// Communication API/CAN/CAN legacy/API/bds_can_getTxBufStatus
///This function returns the status of the Tx buffer of a CAN channel.
///
///=======
/// Remarks:
///=======
///    + Status = number of CAN messages in Tx buffer which have to be sent.
///    + The |GVL_can| is given for usage of defines.
///
///==================================================================		  			===================================================================================================
///Return value    								  									Description
///==================================================================		  			===================================================================================================
///>0																					Number of CAN messages in Tx buffer of the specified CAN channel which have to be sent.
///0																					Tx buffer is empty.
///-1																					Invalid CAN channel.
///5: BDS_CAN_FFI_ACCESS_ERROR_DU16														FFI API access error.
///
///==================================================================		   			===================================================================================================
///
///----------
/// FFI:
///----------
///This API can be used in trusted partitions. For untrusted partitions use |bds_can_getTxBufStatus_ffi|. See Freedom from Interference (FFI) concept for more details.
///
///=======
///Code Example:
///=======
///============================================================================
///
///PROGRAM appl_Task_1
///  VAR
///  
///    numMsg_s32: DINT := 16#00;
///  END_VAR
/// 
///  numMsg_s32 := bds_can_getTxBufStatus(BDS_CAN_1_D);
/// 
///  IF (numMsg_s32 > 0) THEN
///  
///    (* TX buffer contains still messages which could not be sent. If CAN channel
///       is in operational mode the messages will be sent as soon as possible. *)
///	   
///  END_IF
///END
///
///============================================================================
{attribute 'external_name' := 'cmp_rts_bds_can_getTxBufStatus'}
FUNCTION bds_can_getTxBufStatus : DINT
VAR_INPUT
	///Indicates the CAN channel.Possible values are
	///    + BDS_CAN_1_D(0)
	///    + BDS_CAN_2_D(1)
	///    + BDS_CAN_3_D(2)
	///	+ BDS_CAN_4_D(3)
	chnl_e: bds_can_Chnl_te;
END_VAR

END_FUNCTION

// Communication API/CAN/CAN_FFI_API/bds_can_getTxBufStatus_ffi
{attribute 'external_name' := 'cmp_rts_bds_can_getTxBufStatus_ffi'}
FUNCTION bds_can_getTxBufStatus_ffi : DINT
VAR_INPUT
	///Indicates the CAN channel.Possible values are
	///    + BDS_CAN_1_D(0)
	///    + BDS_CAN_2_D(1)
	///    + BDS_CAN_3_D(2)
	///	+ BDS_CAN_4_D(3)
	chnl_e: bds_can_Chnl_te;
END_VAR

END_FUNCTION

// Communication API/CAN/CAN legacy/API/bds_can_initTxDatabox
///This function initializes a CAN transmit databox.
///
///=======
/// Remarks:
///=======
///    + The use of transmit databoxes is optional!
///    + The transmit databoxes must be defined by easyConfig before using this function.
///    + Each transmit databox has to be initialized before it can be used!
///    + If a transmit databox is initialized already it can be inititalized again with new parameters. But if there is a pending message in this transmit databox it will be not sent because the databox is cleared during the initialization.
///    + The |GVL_can| is given for usage of defines.
///    + This API should be called once in Application
///
///----------
/// FFI:
///----------
///This API can be used in trusted partitions only. See Freedom from Interference (FFI) concept for more details.
///
///==================================================================		  			===================================================================================================
///Return value    								  									Description
///==================================================================		  			===================================================================================================
///0: BDS_CAN_ERR_NO_ERRORS_DU16														Function is called without errors. Transmit databox was initialized successfully.
///9: BDS_CAN_ERR_DATABOXNUM_DU16														Invalid transmit databox number.
///14: BDS_CAN_ERR_CHNL_DU16															Unknown CAN channel.
///15: BDS_CAN_ERR_ID_DU16																Invalid CAN identifier.
///16: BDS_CAN_ERR_FORMAT_DU16															Invalid message format.
///
///==================================================================		   			===================================================================================================
///
///=======
///Code Example:
///=======
///============================================================================
///
///PROGRAM PLC_PRG
///  VAR
///  	flag: BOOL;
///
///	status_u16: UINT;
///
///	DataboxData_au8: ARRAY[1..8] OF USINT;
///
///	free_count: INT;
///
///  END_VAR
///
///  (* remark: number of CAN TX databoxes must be configured in easyConfig *)
///
///  (* initialize Tx data box #1 with standard CAN Id = 16#34 *)
/// 
///IF flag = FALSE THEN
///
///	status_u16 := bds_can_initTxDatabox(BDS_CAN_1_D, 3, 16#34, BDS_CAN_STD_DU8);
///
///	bds_can_init(BDS_CAN_1_D, BDS_BAUD_500K_DU32);
///
///	flag:= TRUE;
///
///END_IF
///  (* ... *)
///END
///
///PROGRAM appl_Task_1
///  VAR
///    DataboxData_au8: ARRAY[1..8] OF USINT;
///  END_VAR
///
///  DataboxData_au8[1] := 5;
///  DataboxData_au8[2] := 7;
///
///  if (0 = bds_can_sendDatabox(BDS_CAN_3_D, 1, 2, DataboxData_au8)) THEN
///    (* ok, message will be sent. *)
///  END_IF
///END
///
///============================================================================
{attribute 'external_name' := 'cmp_rts_bds_can_initTxDatabox'}
FUNCTION bds_can_initTxDatabox : UINT
VAR_INPUT
	///Indicates the CAN channel.Possible values are
	///    + BDS_CAN_1_D(0)
	///    + BDS_CAN_2_D(1)
	///    + BDS_CAN_3_D(2)
	///	+ BDS_CAN_4_D(3)
	chnl_e: bds_can_Chnl_te;
	///Transmit databox number.
	///
	///Each transmit databox is numbered separately for each CAN channel.
	///
	///Value range: 1 .. n.
	///
	///n is the number of databoxes configured by easyConfig. 
	databoxNum_u16: UINT;
	///Identifier of CAN message.
	///
	///Value range:
	///    + 16#000 .. 16#7FF (11-bit standard format)
	///    + 16#00000000 .. 16#1FFFFFFF (29-bit extented format)
	id_u32: UDINT;
	///Indicates the format of the CAN message.
	///
	///Value range:
	///    + BDS_CAN_STD_DU8  (11-bit standard format)
	///    + BDS_CAN_EXD_DU8  (29-bit extented format)
	format_u8: USINT;
END_VAR

END_FUNCTION

// Communication API/CAN/CAN legacy/API/bds_can_sendDatabox
///Sends a message via transmit databox.
///
///=======
/// Remarks:
///=======
///    + The number of required transmit databoxes must be defined by easyConfig.
///    + The specified transmit databox has to be initialized by |bds_can_initTxDatabox| before using this function.
///    + A transmit databox buffers only the actual message.
///    + A message in a transmit databox (which was not sent) can be overwritten by a new order. No error will occur!
///    + Function |bds_can_isTxDataboxFree| can be used in order to check whether a transmit databox is free again.
///    + Messages in transmit data boxes will be sent before messages in transmit buffer (|bds_can_sendData|).
///    + The time interval for sending the messages can be defined with the function |bds_can_setTxDelay|.
///    + The |GVL_can| is given for usage of defines.
///
///----------
/// FFI:
///----------
///This API can be used in trusted partitions. For untrusted partitions use |bds_can_sendDatabox_ffi|. See Freedom from Interference (FFI) concept for more details.
///
///==================================================================		  			===================================================================================================
///Return value    								  									Description
///==================================================================		  			===================================================================================================
///0: BDS_CAN_ERR_NO_ERRORS_DU16														Function is called without errors. CAN message will be sent.
///9: BDS_CAN_ERR_DATABOXNUM_DU16														Invalid transmit databox number.
///14: BDS_CAN_ERR_CHNL_DU16															Unknown CAN channel.
///17: BDS_CAN_ERR_NUM_DATA_DU16														Invalid number of data bytes.
///60: BDS_CAN_ERR_INVALID_ADDR_DU16													Invalid address (parameter data_pau8).
///62: BDS_CAN_ERR_DATABOX_NOINIT_DU16													Transmit databox is not initialized.
///5: BDS_CAN_FFI_ACCESS_ERROR_DU16														FFI API access error.
///
///==================================================================		   			===================================================================================================
///
///=======
///Code Example:
///=======
///============================================================================
///
///PROGRAM PLC_PRG
///  VAR
///  	flag: BOOL;
///
///	status_u16: UINT;
///
///	DataboxData_au8: ARRAY[1..8] OF USINT;
///
///	free_count: INT;
///
///  END_VAR
///
///  (* remark: number of CAN TX databoxes must be configured in easyConfig *)
///
///  (* initialize Tx data box #1 with standard CAN Id = 16#34 *)
/// 
///IF flag = FALSE THEN
///
///	status_u16 := bds_can_initTxDatabox(BDS_CAN_1_D, 3, 16#34, BDS_CAN_STD_DU8);
///
///	bds_can_init(BDS_CAN_3_D, BDS_BAUD_500K_DU32);
///
///	flag:= TRUE;
///
///END_IF
///  (* ... *)
///  
///END
///
///PROGRAM appl_Task_1
///  VAR
///    DataboxData_au8: ARRAY[1..8] OF USINT;
///
///  END_VAR
///
///  DataboxData_au8[1] := 5;
///
///  DataboxData_au8[2] := 7;
///
///  if (0 = bds_can_sendDatabox(BDS_CAN_3_D, 1, 2, DataboxData_au8)) THEN
///  
///    (* ok, message will be sent. *)
///	
///  END_IF
///END
///
///============================================================================
{attribute 'external_name' := 'cmp_rts_bds_can_sendDatabox'}
FUNCTION bds_can_sendDatabox : UINT
VAR_INPUT
	///Indicates the CAN channel.Possible values are
	///    + BDS_CAN_1_D(0)
	///    + BDS_CAN_2_D(1)
	///    + BDS_CAN_3_D(2)
	///	+ BDS_CAN_4_D(3)
	chnl_e: bds_can_Chnl_te;
	///Transmit databox number.
	///
	///Each transmit databox is numbered separately for each CAN channel.
	///
	///Value range: 1 .. n.
	///
	///n is the number of Tx databoxes configured by easyConfig. 
	txDataboxNum_u16: UINT;
	///Number of bytes to be sent.
	///
	///Value range: 0 .. 8
	numBytes_u8: USINT;
	///Pointer to array of data bytes. The number of bytes is contained in parameter numBytes_u8. A NULL pointer is allowed if number of data bytes (parameter numBytes_u8) is zero. 
	data_pau8: POINTER TO USINT;
END_VAR

END_FUNCTION

// Communication API/CAN/CAN legacy/API/bds_can_isTxDataboxFree
///This function checks whether a transmit databox is free again. A transmit databox is free again if it was possible to send the last CAN message via the bus.
///
///=======
/// Remarks:
///=======
///    + The use of transmit databoxes is optional!
///    + The transmit databoxes of that CAN channel has to be defined by easyConfig tool and that transmit databox has to be initialised by bds_can_initTxDatabox before using this function.
///    + This function can be used to prevent overwriting of a message that has not yet been sent in a send databox, by checking whether the previous message was actually sent before writing the new message to the databox.
///    + How quickly a databox is free again for sending greatly depends on the baud rate and the bus load.
///    + The |GVL_can| is given for usage of defines.
///
///----------
/// FFI:
///----------
///This API can be used in trusted partitions. For untrusted partitions use |bds_can_isTxChannelFree_ffi|. See Freedom from Interference (FFI) concept for more details.
///
///==================================================================		  			===================================================================================================
///Return value    								  									Description
///==================================================================		  			===================================================================================================
///0: BDS_CAN_TX_DATABOX_EMPTY_DU16													No error. Databox is empty.
///1: BDS_CAN_TX_DATABOX_NOT_EMPTY_DU16												No error. Databox is not empty.
///9: BDS_CAN_ERR_DATABOXNUM_DU16														Invalid databox number.
///14: BDS_CAN_ERR_CHNL_DU16															Unknown CAN channel.
///62: BDS_CAN_ERR_DATABOX_NOINIT_DU16													Databox is not initialized.
///5: BDS_CAN_FFI_ACCESS_ERROR_DU16														FFI API access error.
///
///==================================================================		   			===================================================================================================
///
///=======
///Code Example:
///=======
///============================================================================
///
///PROGRAM PLC_PRG
///
///  VAR
///  	flag: BOOL;
///
///	status_u16: UINT;
///
///	DataboxData_au8: ARRAY[1..8] OF USINT;
///
///	free_count: INT;
///
///  END_VAR
///
///  (* remark: number of CAN TX databoxes must be configured in easyConfig *)
///
///  (* initialize Tx data box #1 with standard CAN Id = 16#34 *)
/// 
///IF flag = FALSE THEN
///
///	status_u16 := bds_can_initTxDatabox(BDS_CAN_1_D, 3, 16#34, BDS_CAN_STD_DU8);
///
///	bds_can_init(BDS_CAN_1_D, BDS_BAUD_500K_DU32);
///
///	flag:= TRUE;
///
///END_IF
///
///PROGRAM appl_Task_1
///  VAR
///  
///  END_VAR
///
///  IF (0 = bds_can_isTxDataboxFree(BDS_CAN_1_D, 1)) THEN
///  
///    (* transmit databox 1 on CAN channel 1 is free and can be loaded again *)
///    (* ... *)
///	
///  END_IF
///END
///
///============================================================================
{attribute 'external_name' := 'cmp_rts_bds_can_isTxDataboxFree'}
FUNCTION bds_can_isTxDataboxFree : UINT
VAR_INPUT
	///Indicates the CAN channel.Possible values are
	///    + BDS_CAN_1_D(0)
	///    + BDS_CAN_2_D(1)
	///    + BDS_CAN_3_D(2)
	///	+ BDS_CAN_4_D(3)
	chnl_e: bds_can_Chnl_te;
	///Transmit databox number.
	///
	///Each transmit databox is numbered separately for each CAN channel.
	///
	///Value range: 1 .. n.
	///
	///n is the number of databoxes configured by easyConfig. 
	txDataboxNum_u16: UINT;
END_VAR

END_FUNCTION

// Communication API/CAN/CAN_FFI_API/bds_can_isTxChannelFree_ffi
{attribute 'external_name' := 'cmp_rts_bds_can_isTxChannelFree_ffi'}
FUNCTION bds_can_isTxChannelFree_ffi : UINT
VAR_INPUT
	///Indicates the CAN channel.Possible values are
	///    + BDS_CAN_1_D(0)
	///    + BDS_CAN_2_D(1)
	///    + BDS_CAN_3_D(2)
	///	+ BDS_CAN_4_D(3)
	chnl_e: bds_can_Chnl_te;
END_VAR

END_FUNCTION

// Communication API/CAN/CAN legacy/API/bds_can_sendData
///Sends a message via the specified CAN channel.
///
///=======
/// Remarks:
///=======
///    + The CAN channel is not buffered until a buffer is registered within easyConfig.
///    + If a buffer is registered then messages are saved in buffer and will be sent in a background process as fast as possible. The buffer principle is first in first out (FIFO).
///    + The time interval for sending the messages can be defined with the function |bds_can_setTxDelay|.
///    + Messages in transmit data boxes (|bds_can_sendDatabox|) will be sent before messages in transmit buffer (|bds_can_sendData|).
///    + The |GVL_can| is given for usage of defines.
///
///----------
/// FFI:
///----------
///This API can be used in trusted partitions. For untrusted partitions use |bds_can_sendData_ffi|. See Freedom from Interference (FFI) concept for more details.
///
///==================================================================		  			===================================================================================================
///Return value    								  									Description
///==================================================================		  			===================================================================================================
///0: BDS_CAN_ERR_NO_ERRORS_DU16														Function is called without errors. CAN message will be sent.
///14: BDS_CAN_ERR_CHNL_DU16															Unknown CAN channel.
///15: BDS_CAN_ERR_ID_DU16																Invalid CAN identifier.
///16: BDS_CAN_ERR_FORMAT_DU16															Invalid message format.
///17: BDS_CAN_ERR_NUM_DATA_DU16														Invalid number of data bytes.
///20: BDS_CAN_ERR_TXBUF_OVFL_DU16														CAN message could not be sent, because of send buffer is full. *1)
///60: BDS_CAN_ERR_INVALID_ADDR_DU16													Invalid address (parameter data_pau8).
///5: BDS_CAN_FFI_ACCESS_ERROR_DU16														FFI API access error.
///
///==================================================================		   			===================================================================================================
///
///possible reasons:
///    + API
///	    + No can send buffer was registered or buffer registered is too small; see buffer configuration in easyConfig.
///        + To many CAN messages have to be sent per time (more orders exceed performance of sending); use higher baudrate, see bds_can_init()
///        + To many CAN messages have to be sent per time by CAN send databoxes; (sending by databoxes is preferred! see bds_can_sendDatabox()
///        + A TX delay time with bds_can_setTxDelay() is defined, which is too big for the number of messages to be sent.
///    + External factors
///        + CAN bus is busy by CAN messages with higher priorities sending by other ECU's so that CAN messages of the own ECU can not be sent.
///        + The sending of CAN messages is delayed due to CAN BUS error(s). Bus-off states will be recovered automatically.
///
///=======
///Code Example:
///=======
///============================================================================
///
///PROGRAM PLC_PRG
///  VAR
///  
///  END_VAR
///
///  (* remark: a CAN TX buffer must be configured in easyConfig *)
///
///  (* re-initialize can channel 1 with 250KBaud. Call the bds_can_init API once *)
///  
///  bds_can_init(BDS_CAN_1_D, BDS_BAUD_250K_DU32);
///
///  (* ... *)
///  
///END
///
///PROGRAM appl_Task_1
///  VAR
///    data_au8: ARRAY[0..7] OF USINT;
///  END_VAR
///
///  data_au8[0] := 5;
///  data_au8[1] := 7;
///
///  IF (0 = bds_can_sendData(BDS_CAN_1_D, 16#123456, BDS_CAN_EXD_DU8, 2, ADR(data_au8))) THEN
///  
///    (* ok, message is buffered and will be sent as fast as possible. *)
///	
///  END_IF
///END
///
///============================================================================
{attribute 'external_name' := 'cmp_rts_bds_can_sendData'}
FUNCTION bds_can_sendData : UINT
VAR_INPUT
	///Indicates the CAN channel.Possible values are
	///    + BDS_CAN_1_D(0)
	///    + BDS_CAN_2_D(1)
	///    + BDS_CAN_3_D(2)
	///	+ BDS_CAN_4_D(3)
	chnl_e: bds_can_Chnl_te;
	///Identifier of CAN message.
	///
	///Value range:
	///    - 16#000 .. 16#7FF (11-bit standard format)
	///    - 16#00000000 .. 16#1FFFFFFF (29-bit extented format)
	id_u32: UDINT;
	///Indicates the format of the CAN message.
	///
	///Value range:
	///    + BDS_CAN_STD_DU8  (11-bit standard format)
	///    + BDS_CAN_EXD_DU8  (29-bit extented format)
	format_u8: USINT;
	///Number of bytes to be sent.
	///
	///Value range: 0 .. 8
	numBytes_u8: USINT;
	///Pointer to array of data bytes. The number of bytes is contained in parameter numBytes_u8. A NULL pointer is allowed if number of data bytes (parameter numBytes_u8) is zero. 
	data_pau8: POINTER TO USINT;
END_VAR

END_FUNCTION

// Communication API/CAN/CAN legacy/API/bds_can_setTxDelay
///The bds_can_setTxDelay function can be used to define an optional delay time for sending CAN messages.
///
///=======
/// Remarks:
///=======
///    + Without executing this function the default delay time = 0 is used.
///    + A delay time > 0 should be only specified, if another controller is not able to receive the CAN messages with full speed.
///    + For each CAN channel another delay time can be specified.
///    + Only messages which are sent with the functions |bds_can_sendDatabox|, |bds_can_sendData| and all messages of ISOBUS module will be delayed.
///    + Signal based CAN messages, XCP and UDS messages are not impacted by this function.
///    + If an error occurs during execution of this function, the actual delay time will be not modified.
///    + The |GVL_can| is given for usage of defines.
///
///----------
/// FFI:
///----------
///This API can be used in trusted partitions only. See Freedom from Interference (FFI) concept for more details.
///
///==================================================================		  			===================================================================================================
///Return value    								  									Description
///==================================================================		  			===================================================================================================
///0: BDS_CAN_ERR_NO_ERRORS_DU16														Function is called without errors. Message data returned in msg_s are valid.
///14: BDS_CAN_ERR_CHNL_DU16															Unknown CAN channel.
///
///==================================================================		   			===================================================================================================
///
///=======
///Code Example:
///=======
///============================================================================
///
///PROGRAM PLC_PRG
///  VAR
///  
///  END_VAR
///
///  (* set the minimum TX delay time to 2ms for CAN channel 1 *)
///  
///IF flag = FALSE THEN
///
///	  bds_can_setTxDelay(BDS_CAN_1_D, 2);
///
///	flag:= TRUE;
///
///END_IF
///  (* ... *)
///END
///
///============================================================================
{attribute 'external_name' := 'cmp_rts_bds_can_setTxDelay'}
FUNCTION bds_can_setTxDelay : UINT
VAR_INPUT
	///Indicates the CAN channel.Possible values are
	///    + BDS_CAN_1_D(0)
	///    + BDS_CAN_2_D(1)
	///    + BDS_CAN_3_D(2)
	///	+ BDS_CAN_4_D(3)
	chnl_e: bds_can_Chnl_te;
	///Minimum delay time in ms between two sent can messages.
	///
	///Value range: 0 .. 65535.
	///
	///0 = no delay time, means that the can messages will be sent as fast as possible.
	time_u16: UINT;
END_VAR

END_FUNCTION

// Communication API/CAN/CAN_FFI_API/bds_can_sendData_ffi
{attribute 'external_name' := 'cmp_rts_bds_can_sendData_ffi'}
FUNCTION bds_can_sendData_ffi : UINT
VAR_INPUT
	///Indicates the CAN channel.Possible values are
	///    + BDS_CAN_1_D(0)
	///    + BDS_CAN_2_D(1)
	///    + BDS_CAN_3_D(2)
	///	+ BDS_CAN_4_D(3)
	chnl_e: bds_can_Chnl_te;
	///Identifier of CAN message.
	///
	///Value range:
	///    - 16#000 .. 16#7FF (11-bit standard format)
	///    - 16#00000000 .. 16#1FFFFFFF (29-bit extented format)
	id_u32: UDINT;
	///Indicates the format of the CAN message.
	///
	///Value range:
	///    + BDS_CAN_STD_DU8  (11-bit standard format)
	///    + BDS_CAN_EXD_DU8  (29-bit extented format)
	format_u8: USINT;
	///Number of bytes to be sent.
	///
	///Value range: 0 .. 8
	numBytes_u8: USINT;
	///Pointer to array of data bytes. The number of bytes is contained in parameter numBytes_u8. A NULL pointer is allowed if number of data bytes (parameter numBytes_u8) is zero. 
	data_pau8: POINTER TO USINT;
END_VAR

END_FUNCTION

// Communication API/CAN/CAN_FFI_API/bds_can_sendDatabox_ffi
{attribute 'external_name' := 'cmp_rts_bds_can_sendDatabox_ffi'}
FUNCTION bds_can_sendDatabox_ffi : UINT
VAR_INPUT
	///Indicates the CAN channel.Possible values are
	///    + BDS_CAN_1_D(0)
	///    + BDS_CAN_2_D(1)
	///    + BDS_CAN_3_D(2)
	///	+ BDS_CAN_4_D(3)
	chnl_e: bds_can_Chnl_te;
	///Transmit databox number.
	///
	///Each transmit databox is numbered separately for each CAN channel.
	///
	///Value range: 1 .. n.
	///
	///n is the number of Tx databoxes configured by easyConfig. 
	txDataboxNum_u16: UINT;
	///Number of bytes to be sent.
	///
	///Value range: 0 .. 8
	numBytes_u8: USINT;
	///Pointer to array of data bytes. The number of bytes is contained in parameter numBytes_u8. A NULL pointer is allowed if number of data bytes (parameter numBytes_u8) is zero. 
	data_pau8: POINTER TO USINT;
END_VAR

END_FUNCTION

// Communication API/CAN/CAN legacy/API/bds_can_isTxChannelFree
///This function checks whether a complete CAN transmit channel is empty.
///
///=======
/// Remarks:
///=======
///    + Empty means that there is no message to send in hardware CAN controller and in any Tx databox (if registered and initialized) and Tx buffer (if registered) is empty.
///    + This function can be used in order to check if a previous message was sent completely on CAN bus. 
///    + The |GVL_can| is given for usage of defines.
///
///----------
/// FFI:
///----------
///This API can be used in trusted partitions. For untrusted partitions use |bds_can_isTxDataboxFree_ffi|. See Freedom from Interference (FFI) concept for more details.
///
///==================================================================		  			===================================================================================================
///Return value    								  									Description
///==================================================================		  			===================================================================================================
///0: BDS_CAN_TX_CHANNEL_EMPTY_DU16													No error. CAN transmit channel is empty. No CAN message has to be sent at the moment.
///1: BDS_CAN_TX_CHANNEL_NOT_EMPTY_DU16												No error. CAN transmit channel is not empty. Sending of a message is still in progress and/or CAN Tx messages are still buffered for sending. 
///2: BDS_CAN_TX_CHANNEL_INV_CAN_DU16													Unknown CAN channel.
///5: BDS_CAN_FFI_ACCESS_ERROR_DU16														FFI API access error.
///
///==================================================================		   			===================================================================================================
///
///=======
///Code Example:
///=======
///============================================================================
///
///PROGRAM appl_Task_1
///  VAR
///  
///  END_VAR
///
///  IF (BDS_CAN_TX_CHANNEL_EMPTY_DU16 = bds_can_isTxChannelFree(BDS_CAN_1_D)) THEN
///  
///    (* All TX databoxes and TX buffer on CAN channel 1 are empty. *)
///    (* ... *)
///	
///  END_IF
///END
///
///============================================================================
{attribute 'external_name' := 'cmp_rts_bds_can_isTxChannelFree'}
FUNCTION bds_can_isTxChannelFree : UINT
VAR_INPUT
	///Indicates the CAN channel.Possible values are
	///    + BDS_CAN_1_D(0)
	///    + BDS_CAN_2_D(1)
	///    + BDS_CAN_3_D(2)
	///	+ BDS_CAN_4_D(3)
	chnl_e: bds_can_Chnl_te;
END_VAR

END_FUNCTION

// Communication API/CAN/CAN_FFI_API/bds_can_isTxDataboxFree_ffi
{attribute 'external_name' := 'cmp_rts_bds_can_isTxDataboxFree_ffi'}
FUNCTION bds_can_isTxDataboxFree_ffi : UINT
VAR_INPUT
	///Indicates the CAN channel.Possible values are
	///    + BDS_CAN_1_D(0)
	///    + BDS_CAN_2_D(1)
	///    + BDS_CAN_3_D(2)
	///	+ BDS_CAN_4_D(3)
	chnl_e: bds_can_Chnl_te;
	///Transmit databox number.
	///
	///Each transmit databox is numbered separately for each CAN channel.
	///
	///Value range: 1 .. n.
	///
	///n is the number of databoxes configured by easyConfig. 
	txDataboxNum_u16: UINT;
END_VAR

END_FUNCTION

// Communication API/CAN/CAN signal based/API/bds_can_sendSignal
///This function is used to transmit message with signal data specified by signal ID on the CAN bus.
///
///Signals are part of PDU, call to this API would cause the PDU to be sent on bus but with the signal contents updated by the signal data pointer. 
///
///This API is responsible for transmission of PDU (for Tx mode= Direct) and updation of signal data (for Tx mode= Cyclic).
///
///=======
/// Remarks:
///=======
///    + Signals referred here are available upon a valid DBC import. 
///    + The parameters of the signal such as Signal ID, length and signal data pointer are passed as parameters to the function while the CAN ID would correspond to the PDU the signal is mapped to.
///    + Easy Config tool allows import of DBC file and selection of frames and signals for the respective CAN nodes.
///    + Signal and PDU properties like Transmission type, no. of repetitions, signal length and so on shall be configured from easyConfig cloud tool.
///    + Interaction Layer Protocol Data Unit(IPDU - a collection of messages transmitted between nodes in a network. 
///    + A sending node packs the messages into an I-PDU in the Interaction Layer (IL) and then transmits them to the network in the Data Link Layer (DLL). 
///    + A receiving node passes each I-PDU from the DLL and to the IL. There, it unpacks the messages and use their contents in the application.
///    + The |GVL_can| is given for usage of defines.
///    + Signal IDs can be located in the post build configuration file - linCanSignals_easyConfig.xml.
///
///----------
/// FFI:
///----------
///This API can be used in trusted partitions only. See Freedom from Interference (FFI) concept for more details.
///
///----------
/// NOTICE:
///----------
///- For signals imported from dbc file,the signal type information comes from dbc. This would generally be of static types like USINT, UINT, SINT, INT. In order to be able to change the length of signal, it requires that the signal is of type USINT_DYN.
///So, for all signals imported from dbc, the length parameter in API has to be set to 0.
///
///==================================================================		  			===================================================================================================
///Return value    								  									Description
///==================================================================		  			===================================================================================================
///BDS_CAN_ERR_NO_ERRORS_DU16 (= 0)													Signal transmission successful.
///BDS_CANSIG_ERR_TX_FAIL_DU16(=117)													Transmission failure.
///BDS_CANSIG_ERR_TX_NOSERVICE_DU16(=119)												Service not available-PDU inactive.
///BDS_CANSIG_ERR_TX_DATAPTR_DU16(=114)												Invalid data pointer address.
///BDS_CANSIG_ERR_NUM_TX_SIG_DU16(=112)												Invalid Signal ID.
///
///==================================================================		   			===================================================================================================
///
///=======
///Code Example:
///=======
///============================================================================
///
///PROGRAM appl_10ms_task
///  VAR
///  
///    bds_IPduGrpVctr_au8:ARRAY[0..1] OF USINT;
///	
///    signaldata_au8: ARRAY[0..7] OF USINT;
///	
///    length_u16: UINT := 16#00;
///	
///  END_VAR
///
///   (* Set the I-PDU and corresponding groups *)
///   (* PDU ,signal and group Ids are available in post build config files from easyConfig *)
/// 
///   bds_can_setMsgGroup(ADR(bds_IPduGrpVctr_au8),ComConf_ComIPduGroup_ComIPduGroup_C_Tx, 1);
///   
///   bds_can_startAllMsgGroups(ADR(bds_IPduGrpVctr_au8), 1) ;
///
///   IF ( 0 = bds_can_sendSignal(ComConf_ComSignal_ComSignal_C_xTx, ADR(signaldata_au8), length_u16) ) THEN
///   
///     (* ok,message is sent on bus with updated signal data *)
///   END_IF
///END
///
///============================================================================
{attribute 'external_name' := 'cmp_rts_bds_can_sendSignal'}
FUNCTION bds_can_sendSignal : UINT
VAR_INPUT
	///ID of the signal to be sent.
	signalId_u16: UINT;
	///Pointer array to the data to be transmitted.
	signalDataPtr_au8: POINTER TO USINT;
	///No. of bytes of data to be sent (for dynamic type signal)
	///	
	///- 0, for static type signals (imported from dbc, refer NOTICE above)
	length_u16: UINT;
END_VAR

END_FUNCTION

// Communication API/CAN/CAN signal based/API/bds_can_setMsgGroup
///A PDU group contains multiple PDUs and each PDU contains one or more signals.
///
///Every message/PDU should be activated before communication. To do this it is required to activate the PDU group in which it is present. This function sets the PDU group specified by group ID, which has to be enabled later by API |bds_can_startAllMsgGroups|.
///
///   
///=======
/// Remarks:
///=======
///    + PDU and message are the same in this context. When it is said that PDU is active, it also means that the message is active.
///    + PDUs referred here are available upon a valid DBC import. 
///    + With the available resources of RC18-12/40 and RC27-18/40, PDU group: There can be a maximum of 8 PDU groups based on the 4 CAN nodes and for each direction (transmit/receive). When PDUs are imported into CAN nodes on eC by DBC importer, the PDUs are put into respective groups. 
///    + To set a PDU, it is necessary to set the PDU group that contains the PDU. 
///    + This API can be called anywhere in the ASW - at init or inside cyclic task.
///    + The PDU groups are generated when we import DBC or add the frame to the CAN channel from eC.
///    + The PDU group name generated will look like ComConf_ComIPduGroup_ComIPduGroup_CAN "channel number"_TX and  ComConf_ComIPduGroup_ComIPduGroup_CAN "channel number"_RX. 
///    + Example:  For CAN 3 the PDU group will look like "ComConf_ComIPduGroup_ComIPduGroup_CAN_3_TX" and   "ComConf_ComIPduGroup_ComIPduGroup_CAN_3_RX".
///    + Interaction Layer Protocol Data Unit (IPDU) - a collection of messages transmitted between nodes in a network. 
///    + A sending node packs the messages into an I-PDU in the Interaction Layer (IL) and then transmits them to the network in the Data Link Layer (DLL). 
///    + A receiving node passes each I-PDU from the DLL and to the IL. There, it unpacks the messages and use their contents in the application.
///	   + The |GVL_can| is given for usage of defines.
///    + PDU and PDU group IDs can be located in the post build configuration file - linCanSignals_easyConfig.xml.
///
///----------
/// FFI:
///----------
///This API can be used in trusted partitions only. See Freedom from Interference (FFI) concept for more details.
///
///==================================================================		  			===================================================================================================
///Return value    								  									Description
///==================================================================		  			===================================================================================================
///BDS_CAN_ERR_NO_ERRORS_DU16 (= 0)													PDU group setting successful.
///BDS_CANSIG_ERR_NULLIPDUVECTOR_DU16(=110)											Invalid Group vector array address.
///BDS_CANSIG_ERR_BITFLAG_DU16(=111)													Invalid parameter bitval.
///
///==================================================================		   			===================================================================================================
///
///=======
///Code Example:
///=======
///============================================================================
///
///PROGRAM appl_10ms_task
///  VAR
///  
///    bds_IPduGrpVctr_au8:ARRAY[0..1] OF USINT;
///  END_VAR
///
///IF ( 0 = bds_can_setMsgGroup(ADR(bds_IPduGrpVctr_au8),ComConf_ComIPduGroup_ComIPduGroup_CAN_1_Tx, 1) ) THEN
///
///    (* ComIPduGroup_CAN_1_TX PDU group is set successfully *)
///    (* All PDUs of this group is now set, next step is to enable *)
///END_IF
///END
///
///============================================================================
{attribute 'external_name' := 'cmp_rts_bds_can_setMsgGroup'}
FUNCTION bds_can_setMsgGroup : UINT
VAR_INPUT
	///PDU group array containing the activation state (stopped = 0/ started = 1) for all message groups.
	rbr_iPduGrpVctr_au8: POINTER TO ARRAY[0..1] OF USINT;
	///PDU group used to identify the corresponding bit in the message group vector.
	ipduGroupId_u16: UINT;
	///New value of the corresponding bit(set PDU =1; reset PDU=0).
	bitval_u8: USINT;
END_VAR

END_FUNCTION

// Communication API/CAN/CAN signal based/API/bds_can_startAllMsgGroups
///This is the master function responsible for activating or deactivating PDU/message groups.
///
///This function is used to activate all PDU/message groups that were set by |bds_can_setMsgGroup|. 
///
///When a PDU group is activated by means of call to this API, all the PDUs belonging to these groups would be activated and the contained signals would be ready for transmission or reception.
///
///=======
/// Remarks:
///=======
///    + PDU and message are the same in this context. 
///    + PDUs referred here are available upon a valid DBC import. 
///    + It is sufficient to call this API once after setting all the PDU groups using the API  |bds_can_setMsgGroup|.
///    + If suppose |bds_can_setMsgGroup| is called sometime later after |bds_can_startAllMsgGroups|, the new PDU group set is still not active and so, bds_can_startAllMsgGroups() will have to be called again. So, everytime a new PDU group is set, it should be activated with this API.
///    + For cyclic signals, the transmission will start soon after the corresponding message and message group is activated by call to this API, the signal data at this instant would be the signal init value defined in eC. Signal data gets updated when the API |bds_can_sendSignal| is called later.
///    + For direct signals, transmission will happen only upon call to |bds_can_sendSignal|.
///    + Interaction Layer Protocol Data Unit(IPDU) - a collection of messages transmitted between nodes in a network. 
///    + A sending node packs the messages into an I-PDU in the Interaction Layer (IL) and then transmits them to the network in the Data Link Layer (DLL). 
///    + A receiving node passes each I-PDU from the DLL and to the IL. There, it unpacks the messages and use their contents in the application.
///    + The |GVL_can| is given for usage of defines.
///    + PDU and PDU group IDs can be located in the post build configuration file - linCanSignals_easyConfig.xml.
///
///----------
/// FFI:
///----------
///This API can be used in trusted partitions only. See Freedom from Interference (FFI) concept for more details.
///
///==================================================================		  			===================================================================================================
///Return value    								  									Description
///==================================================================		  			===================================================================================================
///BDS_CAN_ERR_NO_ERRORS_DU16 (= 0)													PDU groups activation successful.
///BDS_CANSIG_ERR_NULLIPDUVECTOR_DU16(=110)											Invalid Group vector array address.
///BDS_CANSIG_ERR_BITFLAG_DU16(=111)													Invalid parameter Initialize.
///
///==================================================================		   			===================================================================================================
///
///=======
///Code Example:
///=======
///============================================================================
///
///PROGRAM appl_task_1
///  VAR
///  
///    bds_IPduGrpVctr_au8:ARRAY[0..1] OF USINT;
///  END_VAR
///
///bds_can_setMsgGroup(ADR(bds_IPduGrpVctr_au8),ComConf_ComIPduGroup_ComIPduGroup_CAN_1_Tx, 1);
///
///IF ( 0 = bds_can_startAllMsgGroups(ADR(bds_IPduGrpVctr_au8), 1) ) THEN
///
///  (* PDU groups are active and signals ready for transmission(direct) or signal transmission started(cyclic) *)
///END_IF
///END
///
///============================================================================
{attribute 'external_name' := 'cmp_rts_bds_can_startAllMsgGroups'}
FUNCTION bds_can_startAllMsgGroups : UINT
VAR_INPUT
	///PDU group array containing the activation state (stopped = 0/ started = 1) for all PDU groups.
	rbr_iPduGrpVctr_au8: POINTER TO ARRAY[0..1] OF USINT;
	///flag to request initialization of the PDUs
	///	
	///0 = PDU groups will not be activated
	///
	///1 = PDU groups will be activated
	initialize_u8: USINT;
END_VAR

END_FUNCTION

// Communication API/CAN/CAN signal based/API/bds_can_sendSignalGroup
///This function sends the signal group data on the PDU/message.
///
///=======
/// Remarks:
///=======
///    + Before call to this API, it is necessary to update the signal group with data for every group signal belonging to signal group. This is done by using the API bds_can_setGroupSignalData. This function then sends the contents of shadow buffer on the PDU.
///    + Group signals and Signal groups referred here are available upon a valid DBC import. 
///    + Additionally, modification of signal groups by adding group signals to signal group can be done on easyConfig cloud tool.
///    + The parameter SignalGroup ID is passed as parameter to the function while the CAN ID would correspond to the PDU the signal group is mapped to.
///    + Cloud tool allows import of DBC file and selection of frames and signals for the respective CAN nodes.
///    + Signal and PDU properties like Transmission type, number of repetitions, signal length and so on shall be configured from easyConfig cloud tool.
///    + Interaction Layer Protocol Data Unit (IPDU - a collection of messages transmitted between nodes in a network). 
///    + A sending node packs the messages into an I-PDU in the Interaction Layer (IL) and then transmits them to the network in the Data Link Layer (DLL). 
///    + A receiving node passes each I-PDU from the DLL and to the IL. There, it unpacks the messages and use their contents in the application.
///    + The |GVL_can| is given for usage of defines.
///    + Group Signal IDs can be located in the post build configuration file - linCanSignals_easyConfig.xml.
///
///----------
/// FFI:
///----------
///This API can be used in trusted partitions only. See Freedom from Interference (FFI) concept for more details.
///
///==================================================================		  			===================================================================================================
///Return value    								  									Description
///==================================================================		  			===================================================================================================
///BDS_CAN_ERR_NO_ERRORS_DU16 (= 0)													Transmission successful.
///BDS_CANSIG_ERR_TX_NOSERVICE_DU16(=119)												Service not available-PDU inactive.
///
///==================================================================		   			===================================================================================================
///
///=======
///Code Example:
///=======
///============================================================================
///
///PROGRAM appl_task_1
///  VAR
///  
///    bds_IPduGrpVctr_au8:ARRAY[0..1] OF USINT;
///	
///    signaldata_u64: ULINT := 16#1234;
///  END_VAR
///
///  (* Set the I-PDU and corresponding groups *)
///  (* PDU ,signal and group Ids are available in post build config files from easyConfig *)
/// 
///   bds_can_setMsgGroup(ADR(bds_IPduGrpVctr_au8),ComConf_ComIPduGroup_ComIPduGroup_C_Tx, 1);
///   
///   bds_can_startAllMsgGroups(ADR(bds_IPduGrpVctr_au8), 1) ;
///
///   (* update group signal data *)
///   
///   bds_can_setGroupSignalData(ComConf_ComGroupSignal_ComGroupSignal_Tx, signaldata_u64);
///
///   IF ( 0 = bds_can_sendSignalGroup(ComConf_ComSignalGroup_ComSignalGroup_Tx_1) ) THEN
///   
///     (* ok, message is sent on bus with signalgroup data *)
///   END_IF
///END
///
///============================================================================
{attribute 'external_name' := 'cmp_rts_bds_can_sendSignalGroup'}
FUNCTION bds_can_sendSignalGroup : UINT
VAR_INPUT
	///ID of the signal group to be transmitted.
	signalGroupId_u16: UINT;
END_VAR

END_FUNCTION

// Communication API/CAN/CAN signal based/API/bds_can_setGroupSignalData
///This function updates the group signal with the data referenced by signalData parameter.
///
///The updated data is now stored in a shadow buffer of the signal group.
///
///The entire contents of signal group shadow buffer is transmitted on a message/PDU upon call to API |bds_can_sendSignalGroup|.
///
///=======
/// Remarks:
///=======
///    + Group Signals and Signal groups referred here are available upon a valid DBC import. 
///    + Additionally, modification of signal groups by adding group signals to signal group can be done on easyConfig cloud tool.
///    + Group Signal IDs can be located in the post build configuration file - BODAS API library, bds_rts_ec.xml.
///    + The parameters of the signal such as Group Signal ID and signal data are passed as parameters to the function while the CAN ID would correspond to. 
///    + Interaction Layer Protocol Data Unit (IPDU - a collection of messages transmitted between nodes in a network). 
///    + A sending node packs the messages into an I-PDU in the Interaction Layer (IL) and then transmits them to the network in the Data Link Layer (DLL). 
///    + A receiving node passes each I-PDU from the DLL and to the IL. There, it unpacks the messages and use their contents in the application.
///    + The |GVL_can| is given for usage of defines.
///    + Group Signal IDs can be located in the post build configuration file - linCanSignals_easyConfig.xml.
///
///----------
/// FFI:
///----------
///This API can be used in trusted partitions only. See Freedom from Interference (FFI) concept for more details.
///
///==================================================================		  			===================================================================================================
///Parameter	   								  										Description
///==================================================================		  			===================================================================================================
///groupSignalId_u16																	ID of the group signal to be sent.
///signalData_u64																		Signal data for the specified group signal to be transmitted. Maximum size of data is 64 bits(8bytes).
///
///==================================================================		   			===================================================================================================
///
///=======
///Code Example:
///=======
///============================================================================
///
///PROGRAM appl_10ms_task
///  VAR
///  
///    bds_IPduGrpVctr_au8:ARRAY[0..1] OF USINT;
///	
///    signaldata_u64: ULINT := 16#1234;
///  END_VAR
///
///  (* Set the I-PDU and corresponding groups *)
///  (* PDU ,signal and group Ids are available in post build config files from easyConfig *)
/// 
///   bds_can_setMsgGroup(ADR(bds_IPduGrpVctr_au8),ComConf_ComIPduGroup_ComIPduGroup_C_Tx, 1);
///   
///   bds_can_startAllMsgGroups(ADR(bds_IPduGrpVctr_au8), 1) ;
///
///   (* update group signal data *)
///   
///   bds_can_setGroupSignalData(ComConf_ComGroupSignal_ComGroupSignal_Tx, signaldata_u64);
///END
///
///============================================================================
{attribute 'external_name' := 'cmp_rts_bds_can_setGroupSignalData'}
FUNCTION bds_can_setGroupSignalData : BOOL
VAR_INPUT
	///ID of the group signal to be sent.
	groupSignalId_u16: UINT;
	///Signal data for the specified group signal to be transmitted. Maximum size of data is 64 bits(8bytes).
	signalData_u64: ULINT;
END_VAR

END_FUNCTION

// Communication API/CAN/CAN signal based/API/bds_can_receiveSignal
///Signals are part of PDU/message, call to this API would cause the signal data of the PDU/message received on bus to be copied to application defined buffer.
///
///=======
/// Remarks:
///=======
///    + Signals referred here are available upon a valid DBC import. 
///    + The parameters of the signal such as Signal ID, length and signal data pointer are passed as parameters to the function while the CAN ID would correspond to the PDU, the signal is mapped to.
///    + Easy Config tool allows import of DBC file and selection of frames and signals for the respective CAN nodes.
///    + Signal and PDU properties like Transmission type, no. of repetitions, signal length and so on shall be configured from easyConfig cloud tool.
///    + Interaction Layer Protocol Data Unit (IPDU - a collection of messages transmitted between nodes in a network). 
///    + A sending node packs the messages into an I-PDU in the Interaction Layer (IL) and then transmits them to the network in the Data Link Layer (DLL). 
///    + A receiving node passes each I-PDU from the DLL and to the IL. There, it unpacks the messages and use their contents in the application.
///    + The |GVL_can| is given for usage of defines.
///    + Signal IDs can be located in the post build configuration file - linCanSignals_easyConfig.xml.
///
///----------
/// FFI:
///----------
///This API can be used in trusted partitions only. See Freedom from Interference (FFI) concept for more details.
///
///----------
/// NOTICE:
///----------
///The length parameter specifies the no. of bytes of data to be received and it is important to specify exactly the no. of incoming bytes else it would result in length validation failure.
///- For signals imported from dbc file,the signal type information comes from dbc. This would generally be of static types like USINT, UINT, SINT, INT.
///
///==================================================================		  			===================================================================================================
///Return value    								  									Description
///==================================================================		  			===================================================================================================
///BDS_CAN_ERR_NO_ERRORS_DU16 (= 0)													Signal reception successful.
///BDS_CANSIG_ERR_RX_FAIL_DU16(=118)													Reception failure.
///BDS_CANSIG_ERR_RX_NOSERVICE_DU16(=120)												Service not available-PDU inactive.
///BDS_CANSIG_ERR_RX_LENPTR_DU16(=116)													Invalid parameter length.
///BDS_CANSIG_ERR_RX_DATAPTR_DU16(=115)												Invalid data pointer address.
///BDS_CANSIG_ERR_NUM_RX_SIG_DU16(=113)												Invalid Signal ID.
///
///==================================================================		   			===================================================================================================
///
///=======
///Code Example:
///=======
///============================================================================
///
///PROGRAM appl_10ms_task
///  VAR
///    bds_IPduGrpVctr_au8:ARRAY[0..1] OF USINT;
///	
///    Rx_data_au8: ARRAY[0..7] OF USINT;
///	
///    length_u16: UINT := 16#00;
///  END_VAR
///
///  (* Set the I-PDU and corresponding groups *)
///  (* PDU ,signal and group Ids are available in post build config files from easyConfig *)
/// 
///   bds_can_setMsgGroup(ADR(bds_IPduGrpVctr_au8),ComConf_ComIPduGroup_ComIPduGroup_C_Rx, 1);
///   
///   bds_can_startAllMsgGroups(ADR(bds_IPduGrpVctr_au8), 1) ;
///
///   IF ( 0 = bds_can_receiveSignal(ComConf_ComSignal_ComSignal_C_xRx,ADR(Rx_data_au8),length_u16) ) THEN
///   
///     (* Data is stored in Rx_data_au8 *)
///	 
///   END_IF
///END
///
///============================================================================
{attribute 'external_name' := 'cmp_rts_bds_can_receiveSignal'}
FUNCTION bds_can_receiveSignal : UINT
VAR_INPUT
	///ID of the signal to be received.
	signalId_u16: UINT;
	///Pointer array to location where the received signal data shall be stored.
	signalDataPtr_au8: POINTER TO USINT;
	///- No. of bytes of data expected to be received (for dynamic type signal)
	///	
	///- 0 , for static signals(imported from dbc, refer NOTICE above)
	length_u16: UINT;
END_VAR

END_FUNCTION

// Communication API/CAN/CAN signal based/API/bds_can_receiveSignalGroup
///This function copies the contents of a group signal from the received message into the referenced data buffer.
///
///=======
/// Remarks:
///=======
///    + Group Signals and Signal groups referred here are available upon a valid DBC import. 
///    + Additionally, modification of signal groups by adding group signals to signal group can be done on easyConfig cloud tool.
///    + The parameters of the signal such as Group Signal ID, Signal Group ID and signal dataptr are passed as parameters to the function while the CAN ID would correspond to the PDU the signal and signal group is mapped to.
///    + Cloud tool allows import of DBC file and selection of frames and signals for the respective CAN nodes.
///    + Interaction Layer Protocol Data Unit(IPDU - a collection of messages transmitted between nodes in a network. 
///    + A sending node packs the messages into an I-PDU in the Interaction Layer (IL) and then transmits them to the network in the Data Link Layer (DLL). 
///    + A receiving node passes each I-PDU from the DLL and to the IL. There, it unpacks the messages and use their contents in the application.
///    + The |GVL_can| is given for usage of defines.
///    + Group Signal IDs can be located in the post build configuration file - linCanSignals_easyConfig.xml.
///
///----------
/// FFI:
///----------
///This API can be used in trusted partitions only. See Freedom from Interference (FFI) concept for more details.
///
///==================================================================		  			===================================================================================================
///Return value    								  									Description
///==================================================================		  			===================================================================================================
///BDS_CAN_ERR_NO_ERRORS_DU16 (= 0)													Signal Reception successful.
///BDS_CANSIG_ERR_RX_DATAPTR_DU16(=115)												Invalid data pointer address.
///BDS_CANSIG_ERR_RX_NOSERVICE_DU16(=120)												Service not available-PDU inactive.
///
///==================================================================		   			===================================================================================================
///
///=======
///Code Example:
///=======
///============================================================================
///
///PROGRAM appl_task_1
///  VAR
///  
///    bds_IPduGrpVctr_au8:ARRAY[0..1] OF USINT;
///	
///    Rx_data_au8: ARRAY[0..7] OF USINT;
///	
///  END_VAR
///
///  (* Set the I-PDU and corresponding groups *)
///  (* PDU ,signal and group Ids are available in post build config files from easyConfig *)
/// 
///   bds_can_setMsgGroup(ADR(bds_IPduGrpVctr_au8),ComConf_ComIPduGroup_ComIPduGroup_C_Rx, 1);
///   
///   bds_can_startAllMsgGroups(ADR(bds_IPduGrpVctr_au8), 1) ;
///
///   IF ( 0 = bds_can_receiveSignalGroup(ComConf_ComSignalGroup_ComSignalGroup_Rx_1, ComConf_ComGroupSignal_ComGroupSignal_Rx, ADR(Rx_data_au8) ) THEN
///   
///     (* Data is stored in Rx_data_au8 *)
///	 
///   END_IF
///END
///
///============================================================================
{attribute 'external_name' := 'cmp_rts_bds_can_receiveSignalGroup'}
FUNCTION bds_can_receiveSignalGroup : UINT
VAR_INPUT
	///ID of the signal group to be received.
	signalGroupId_u16: UINT;
	///ID of the group signal to be received.
	groupSignalId_u16: UINT;
	///Buffer to which the Group signal data is copied.
	RxDataPtr_au8: POINTER TO BOOL;
END_VAR

END_FUNCTION

// Communication API/CAN/CAN signal based/API/bds_can_resetAllMsgGroups
///This API is used to clear the PDU/message group setting.
///
///This function sets all bits of PDU group entry in the PDU group array to zero.The purpose of this function is to reset all PDUs and PDU groups.
///
///=======
/// Remarks:
///=======
///    + PDU and message are the same in this context. 
///    + PDUs referred here are available upon a valid DBC import.
///    + This API works together with  |bds_can_setMsgGroup|. All the PDU groups that were set from the API |bds_can_setMsgGroup| would be reset to 0. 
///    + This API does not deactivate PDUs. But can be used together with |bds_can_startAllMsgGroups| to deactivate PDUs.
///    + Interaction Layer Protocol Data Unit (IPDU) - a collection of messages transmitted between nodes in a network. 
///    + A sending node packs the messages into an I-PDU in the Interaction Layer (IL) and then transmits them to the network in the Data Link Layer (DLL). 
///    + A receiving node passes each I-PDU from the DLL and to the IL. There, it unpacks the messages and use their contents in the application.
///    + The |GVL_can| is given for usage of defines.
///    + PDU and PDU group IDs can be located in the post build configuration file - linCanSignals_easyConfig.xml.
///
///----------
/// FFI:
///----------
///This API can be used in trusted partitions only. See Freedom from Interference (FFI) concept for more details.
///
///==================================================================		  			===================================================================================================
///Return value    								  									Description
///==================================================================		  			===================================================================================================
///BDS_CAN_ERR_NO_ERRORS_DU16 (= 0)													PDU group reset successful.
///BDS_CANSIG_ERR_NULLIPDUVECTOR_DU16(=110)											Invalid Group vector array address.
///
///==================================================================		   			===================================================================================================
///
///=======
///Code Example:
///=======
///============================================================================
///
///PROGRAM appl_task_1
///  VAR
///  
///    bds_IPduGrpVctr_au8:ARRAY[0..1] OF USINT;
///  END_VAR
///
///IF ( 0 = bds_can_resetAllMsgGroups(ADR(bds_IPduGrpVctr_au8)) ) THEN
///
///  (* All PDU groups reset successfully.Call bds_can_startAllMsgGroups with flag = 0 to deactivate all groups*)
///  
///END_IF
///END
///
///============================================================================
{attribute 'external_name' := 'cmp_rts_bds_can_resetAllMsgGroups'}
FUNCTION bds_can_resetAllMsgGroups : UINT
VAR_INPUT
	///PDU group array containing the activation state (stopped = 0/ started = 1) for all PDU groups.
	rbr_iPduGrpVctr_au8: POINTER TO ARRAY[0..1] OF USINT;
END_VAR

END_FUNCTION

// System API/DSM/API/bds_dsm_delError
///This function resets the status of specific DFC as well as deletes the related DFES entry if it exists. 
///
///=======
/// Remarks:
///=======
///    + The |GVL_dsm| is given for usage of defines.
///
///----------
/// FFI:
///----------
///This API can be used in trusted partitions only. See Freedom from Interference (FFI) concept for more details.
///
///==================================================================		  			===================================================================================================
///Return value    								  									Description
///==================================================================		  			===================================================================================================
///16#0000: BDS_DSM_NO_ERROR_DU16														Both DFES entry and DFC status bit are cleared in DFC status memory.
///16#0001: BDS_DSM_DFC_ERROR_DU16														Invalid DFC.
///16#0009: BDS_DSM_DFC_NOEXIST_DU16													DFC does not exist in DFES.Possible causes:
///																					   + DFC is configured that it is never saved in DFES.
///																					   + DFC is configured to save in DFES but it can not be saved in DFES because DFES is full.
///
///==================================================================		   			===================================================================================================
///=======
///Code Example:
///=======
///============================================================================
///
///PROGRAM BDS_DSM_DEL_ERROR_TEST
///
///VAR
///
///	dfc_s: bds_dsm_dfc_ts;	
///
///	(*Application Error to be deleted*)
///	
///	dfc_ts : DFC_bds_NoDebFault1;
///
///	status_u16: UINT;
///
///END_VAR
///
///dfc_s.id := dfc_ts.DFCid;
///
///(*Deletes the Error status from DFC and related DFES entry*)
///
///status_u16 := bds_dsm_delError(dfc_s); 
///
///if status_u16 = BDS_DSM_NO_ERROR_DU16 THEN
///
///	(*Error has been deleted successfully*)
///
///END_IF
///
///
///============================================================================
///
///
{attribute 'external_name' := 'cmp_rts_bds_dsm_delError'}
FUNCTION bds_dsm_delError : UINT
VAR_INPUT
	///DFC name (identifier) : It is configured using easyConfig tool.
	dfc_s: bds_dsm_dfc_ts;
END_VAR

END_FUNCTION

// System API/DSM/API/bds_dsm_delErrors
///This function is used to reset the status of all DFCs specified by the mask as well as to delete the related DFES entries if they exist.  
///
///=======
/// Remarks:
///=======
///    + The |GVL_dsm| is given for usage of defines.
///
///----------
/// FFI:
///----------
///This API can be used in trusted partitions only. See Freedom from Interference (FFI) concept for more details.
///
///==================================================================		  			===================================================================================================
///Return value    								  									Description
///==================================================================		  			===================================================================================================
///16#0000: BDS_DSM_NO_ERROR_DU16														Update Number of Error is successful.
///16#0005: BDS_DSM_MASK_ERROR_DU16													Invalid Mask.
///
///==================================================================		   			===================================================================================================
///
///
///=======
///Code Example:
///=======
///============================================================================
///
///PROGRAM BDS_DSM_DEL_ERRORS_TEST
///
///VAR
///
///	dfc_s: bds_dsm_dfc_ts;	
///
///	(*Application Error to be deleted*)
///	
///	dfc_ts : DFC_bds_NoDebFault1;
///
///	status_u16: UINT;
///
///END_VAR
///
///dfc_s.id := dfc_ts.DFCid;
///
///(*delete errors according the Mask*)
///
///status_u16 := bds_dsm_delError(BDS_DSM_SET_TESTED_OK_MASK_DU16); 
///
///if status_u16 = BDS_DSM_NO_ERROR_DU16 THEN
///
///	(*Error has been deleted successfully*)
///
///END_IF
///
///
///============================================================================
///
{attribute 'external_name' := 'cmp_rts_bds_dsm_delErrors'}
FUNCTION bds_dsm_delErrors : UINT
VAR_INPUT
	///The kind of error status can be specified in detail by means of this mask.
	///
	///Possible values:
	///    + BDS_DSM_SET_ACTIVE_ERROR_MASK_DU16 (16#18) - Fault is active.
	///    + BDS_DSM_SET_TESTED_ONCE_MASK_DU16 (16#08) - DFC was tested at least once since start or reset.
	///    + BDS_DSM_SET_TESTED_OK_MASK_DU16 (16#20) - DFC was at least once ok tested since start or reset.  
	///    + BDS_DSM_SET_FAILED_SINCE_CLEAR_MASK_DU16 (16#80) - Fault occurred at least once since error was deleted from memory.
	mask_s: UINT;
END_VAR

END_FUNCTION

// I/O API/OUT_LEGACY/bds_out_do_resetError
///Resets an error and unlocks the digital output
///
///=======
/// Remarks:
///=======
///   + After a fault the output is locked but the set point is still valid. With the error is reset, output is also unlocked.
///   + After a hot short circuit the unlock of the power output is only possible after a reactivation time of 2s.
///
///----------
/// FFI:
///----------
///This API can be used in trusted partitions only. See Freedom from Interference (FFI) concept for more details.
///
///==================================================================		  			===================================================================================================
///Return value    								  									Description
///==================================================================		  			===================================================================================================
///0																					No error
///1																					A parameter is invalid.
///2																					Reset not possible (output is locked by MO Module).
///3																					Reactivation time not elapsed.
///
///==================================================================		   			===================================================================================================
///
///=======
///Code Example:
///=======
///============================================================================
///
///PROGRAM appl_10ms_task
///
///VAR
///
///return_u8: USINT := 16#00;
///
///END_VAR
///
///
///
///(* reset error of output K12 *)
///
///return_u8 = bds_out_do_resetError(bds_out_do_signal_te.K12);
///
///
///============================================================================
{attribute 'external_name' := 'cmp_rts_bds_out_do_resetError'}
FUNCTION bds_out_do_resetError : USINT
VAR_INPUT
	///The connector assigned signal name of the output.
	signal_e: UINT;
END_VAR

END_FUNCTION

// I/O API/OUT_LEGACY/bds_out_do_unlock
///Unlocks digital output if there are no errors anymore.
///
///=======
/// Remarks:
///=======
///   + After a fault the output is locked but the set point is still valid.
///   + It is possible to poll the status of the fault. If the error has been healed, then the output can be unlocked.
///   + After a hot short circuit and over current the unlocking of the power output is only possible after a reactivation time of 2s.
///   + For over current fault: After unlocking, the output has to be switched on again using the API. ( see |bds_out_do|)
///
///----------
/// FFI:
///----------
///This API can be used in trusted partitions only. See Freedom from Interference (FFI) concept for more details.
///
///==================================================================		  			===================================================================================================
///Return value    								  									Description
///==================================================================		  			===================================================================================================
///16#0000																				No error, unlocked successfully.
///16#0001																				Error output was locked by the MO Module.
///16#0002																				Error reactivation time not elapsed
///16#0004																				Error DFC_SCB is set.
///16#0008																				Error DFC_SCG is set
///16#0010																				Error DFC_OL is set
///16#0020																				Error DFC_OT is set
///16#0040																				-
///16#0080																				Error OC is reset, output is unlocked
///16#8000																				Error signal is out of range
///
///==================================================================		   			===================================================================================================
///
///=======
///Code Example:
///=======
///============================================================================
///
///PROGRAM appl_10ms_task
///
///VAR
///
///return_u16: UINT := 16#00;
///
///END_VAR
///
///
///
///(* reset error of output K12 *)
///
///return_u16 = bds_out_do_unlock(bds_out_do_signal_te.K12);
///
///
///============================================================================
{attribute 'external_name' := 'cmp_rts_bds_out_do_unlock'}
FUNCTION bds_out_do_unlock : UINT
VAR_INPUT
	///The connector assigned signal name of the output.
	signal_e: UINT;
END_VAR

END_FUNCTION

// I/O API/OUT_LEGACY/bds_out_do
///Sets the digital output to a particular state.
///
///=======
/// Remarks:
///=======
///   + For more information see |bds_out_do_getStatus| and |bds_out_do_resetError|.
///   + This function should be called only once in the application.
///   
///
///----------
/// FFI:
///----------
///This API can be used in trusted partitions . For untrusted partitions use |bds_out_do_ffi|. See Freedom from Interference (FFI) concept for more details.
///
///==================================================================		  			===================================================================================================
///Return value    								  									Description
///==================================================================		  			===================================================================================================
///0																					No error
///1																					Invalid parameter
///2																					Function call was erroneous.
///3																					Output is disabled.
///4																					Output is locked
///5																					Already configured as SAFOUT channel
///
///==================================================================		   			===================================================================================================
///
///=======
///Code Example:
///=======
///============================================================================
///
///PROGRAM PLC_PRG
///
///VAR
///
///	Init_flag_u8:USINT:=0;
///
///END_VAR
///  
///IF(Init_flag_u8=0) THEN (*To make api call once in application*)
///
///	(* activate output K12 *)
///	
///	bds_out_do(bds_out_do_signal_te.K12, STD_ACTIVE);
///	
///	Init_flag_u8:=1;
///  
///END_IF
///
///============================================================================
{attribute 'external_name' := 'cmp_rts_bds_out_do'}
FUNCTION bds_out_do : USINT
VAR_INPUT
	///The connector assigned signal name of the output.
	signal_e: UINT;
	///State of the output.
	///   + STD_IDLE
	///   + STD_ACTIVE
	state_u8: USINT;
END_VAR

END_FUNCTION

// I/O API/OUT_LEGACY/bds_out_do_getStatus
///Provides the status of a digital output.
///
///=======
/// Remarks:
///=======
///   + The status data holds all relevant information of the digital output.
///	   + Part of the status data is also the fault status of every DFC (e.g. stDFC_SCB_u16). 
///
///----------
/// FFI:
///----------
///This API can be used in trusted partitions . For untrusted partitions use |bds_out_do_getStatus_ffi|. See Freedom from Interference (FFI) concept for more details.
///
///==================================================================		  			===================================================================================================
///Return value    								  									Description
///==================================================================		  			===================================================================================================
///0																					No error
///1																					A parameter is invalid.
///
///==================================================================		   			===================================================================================================
///
///=======
///Code Example:
///=======
///============================================================================
///
///PROGRAM appl_10ms_task
///
///VAR
///
///	stK12_s: bds_out_do_ts;
///	
///	ldf_u8: USINT := 16#00;
///
///END_VAR
///
///
///
///(* get the status of output K12 *)
///
///bds_out_do_getStatus(bds_out_do_signal_te.K12, ADR(stK12_s));
///
///
///
///(* get last debounced fault *)
///
///ldf_u8 := bds_dsm_DFC_ldf(stK12_s.stDFC_SCB_u16);
///
///============================================================================
{attribute 'external_name' := 'cmp_rts_bds_out_do_getStatus'}
FUNCTION bds_out_do_getStatus : USINT
VAR_INPUT
	///The connector assigned signal name of the output.
	signal_e: UINT;
	///Storage address of the data.
	data_ps: POINTER TO bds_out_do_ts;
END_VAR

END_FUNCTION

// I/O API/OUT/FFI_API/bds_out_do_getStatus_ffi
{attribute 'external_name' := 'cmp_rts_bds_out_do_getStatus_ffi'}
FUNCTION bds_out_do_getStatus_ffi : USINT
VAR_INPUT
	///The connector assigned signal name of the output.
	signal_e: UINT;
	///Storage address of the data.
	data_ps: POINTER TO bds_out_do_ts;
END_VAR

END_FUNCTION

// System API/DSM/API/Macro Functions/bds_dsm_DFC_ldf
///It returns the last debounced fault bit fields from DFC status word
{attribute 'external_name' := 'cmp_rts_bds_dsm_DFC_ldf'}
FUNCTION bds_dsm_DFC_ldf : USINT
VAR_INPUT
	dfc_u16: UINT;
END_VAR

END_FUNCTION

// I/O API/OUT/FFI_API/bds_out_do_ffi
{attribute 'external_name' := 'cmp_rts_bds_out_do_ffi'}
FUNCTION bds_out_do_ffi : USINT
VAR_INPUT
	///The connector assigned signal name of the output.
	signal_e: UINT;
	///State of the output.
	///   + STD_IDLE
	///   + STD_ACTIVE
	state_u8: USINT;
END_VAR

END_FUNCTION

// I/O API/OUT_LEGACY/bds_out_po
///Sets the proportional output to the given duty cycle.
///
///=======
/// Remarks:
///=======
///   + For more information see |bds_out_po_getStatus| and |bds_out_po_resetError|.
///
///----------
/// FFI:
///----------
///This API can be used in trusted partitions.  For untrusted partitions use |bds_out_po_ffi|. See Freedom from Interference (FFI) concept for more details.
///
///==================================================================		  			===================================================================================================
///Return value    								  									Description
///==================================================================		  			===================================================================================================
///0																					No error.
///1																					A parameter is invalid.
///2																					Function call was erroneous.
///3																					Already configured as POC.
///4																					Output is disabled.
///5																					Output is locked
///6																					Already configured as SAFOUT channel
///
///==================================================================		   			===================================================================================================
///
///=======
///Code Example:
///=======
///============================================================================
///
///PROGRAM appl_10ms_task
///
///VAR
///
///END_VAR
///
///
///(* set a duty cycle of 50% *)
///
///bds_out_po(bds_out_po_signal_te.K73, 500);
///
///============================================================================
{attribute 'external_name' := 'cmp_rts_bds_out_po'}
FUNCTION bds_out_po : USINT
VAR_INPUT
	///The connector assigned signal name of the output.
	signal_e: UINT;
	///Duty cycle [0,1%]
	///   + Range:0 to 1000 
	dc_u16: UINT;
END_VAR

END_FUNCTION

// I/O API/OUT_LEGACY/bds_out_po_getStatus
///Provides the status of the proportional output.
///
///=======
/// Remarks:
///=======
///   + The status data holds all relevant information of the proportional output, see example below.
///   + Part of the status data is also the fault status of every DFC (e.g. stDFC_SCB_u16).
///   + With the macros (e.g. bds_dsm_DFC_ldf) defined in bds_dsm_api.h , respective bit fields of the fault status can be read.
///
///----------
/// FFI:
///----------
///This API can be used in trusted partitions . For untrusted partitions use |bds_out_po_getStatus_ffi|. See Freedom from Interference (FFI) concept for more details.
///
///==================================================================		  			===================================================================================================
///Return value    								  									Description
///==================================================================		  			===================================================================================================
///0																					No error.
///1																					A parameter is invalid.
///
///==================================================================		   			===================================================================================================
///
///=======
///Code Example:
///=======
///============================================================================
///
///PROGRAM appl_10ms_task
///
///VAR
///
///	stK73_s: bds_out_po_ts;
///
///	ldf_u8: USINT := 16#00;
///
///END_VAR
///
///
///
///(* get the status of output K73 *)
///
///bds_out_po_getStatus(bds_out_po_signal_te.K73, ADR(stK73_s));
///
///
///
///(* get last debounced fault *)
///
///ldf_u8 = bds_dsm_DFC_ldf(stK73_s.stDFC_SCB_u16);
///
///
///============================================================================
{attribute 'external_name' := 'cmp_rts_bds_out_po_getStatus'}
FUNCTION bds_out_po_getStatus : USINT
VAR_INPUT
	///The connector assigned signal name of the output.
	signal_e: UINT;
	///Storage address of the data.
	data_ps: POINTER TO bds_out_po_ts;
END_VAR

END_FUNCTION

// I/O API/OUT/FFI_API/bds_out_po_getStatus_ffi
{attribute 'external_name' := 'cmp_rts_bds_out_po_getStatus_ffi'}
FUNCTION bds_out_po_getStatus_ffi : USINT
VAR_INPUT
	///The connector assigned signal name of the output.
	signal_e: UINT;
	///Storage address of the data.
	data_ps: POINTER TO bds_out_po_ts;
END_VAR

END_FUNCTION

// I/O API/OUT_LEGACY/bds_out_po_resetError
///Resets an error and unlocks the proportional output.
///
///=======
/// Remarks:
///=======
///
///   + After a fault, the output is locked but the set point is still valid. With the reset of the error the output is also unlocked.
///   + After a hot short circuit, the unlocking of the power output is only possible after a reactivation time of 2s.
///
///----------
/// FFI:
///----------
///This API can be used in trusted partitions only. See Freedom from Interference (FFI) concept for more details.
///
///==================================================================		  			===================================================================================================
///Return value    								  									Description
///==================================================================		  			===================================================================================================
///0																					No error.
///1																					A parameter is invalid.
///2																					Reset not possible (output is locked by MO Module).
///3																					Reactivation time not elapsed.
///
///==================================================================		   			===================================================================================================
///
///=======
///Code Example:
///=======
///============================================================================
///
///PROGRAM appl_10ms_task
///
///VAR
///
/// return_u8: USINT := 16#00;
///
///END_VAR
///
///
///
///(* reset error of output K73 *)
///
///return_u8 = bds_out_po_resetError(bds_out_po_signal_te.K73);
///
///============================================================================
{attribute 'external_name' := 'cmp_rts_bds_out_po_resetError'}
FUNCTION bds_out_po_resetError : USINT
VAR_INPUT
	///The connector assigned signal name of the output.
	signal_e: UINT;
END_VAR

END_FUNCTION

// I/O API/OUT/FFI_API/bds_out_po_ffi
{attribute 'external_name' := 'cmp_rts_bds_out_po_ffi'}
FUNCTION bds_out_po_ffi : USINT
VAR_INPUT
	///The connector assigned signal name of the output.
	signal_e: UINT;
	///Duty cycle [0,1%]
	///   + Range:0 to 1000 
	dc_u16: UINT;
END_VAR

END_FUNCTION

// I/O API/OUT_LEGACY/bds_out_poc
///Sets the proportional output with current control to a given set point.
///
///=======
/// Remarks:
///=======
///   + A deviation to the set point can be configured with |bds_out_poc_cfg|.
///   + For more information see |bds_out_po_getStatus| and |bds_out_po_resetError|.
///
///----------
/// FFI:
///----------
///This API can be used in trusted partitions . For untrusted partitions use |bds_out_poc_ffi|. See Freedom from Interference (FFI) concept for more details.
///
///------
/// Info:
///------
///
///It is mandatory that the proportional output is configured as proportional output with current control (POC).( see |bds_out_po_cfg|.)
///
///==================================================================		  			===================================================================================================
///Return value    								  									Description
///==================================================================		  			===================================================================================================
///0																					No error.
///1																					A parameter is invalid.
///2																					Not configured as POC.
///3																					Request current out of range.
///4																					Output is disabled.
///5																					Output is locked
///6																					Already configured as SAFOUT channel
///
///==================================================================		   			===================================================================================================
///
///=======
///Code Example:
///=======
///============================================================================
///
///PROGRAM appl_10ms_task
///
///VAR
///
///END_VAR
///
///
///
///(* set a current of 500mA *)
///
///bds_out_poc(bds_out_po_signal_te.K73, 500);
///
///============================================================================
{attribute 'external_name' := 'cmp_rts_bds_out_poc'}
FUNCTION bds_out_poc : USINT
VAR_INPUT
	///The connector assigned signal name of the output.
	signal_e: UINT;
	///Set point [mA].
	///   + Range:0 to 3000/4000. Current control upper limit depends on the used output.
	iSet_u16: UINT;
END_VAR

END_FUNCTION

// I/O API/OUT_LEGACY/bds_out_poc_cfg
///For a proportional output with current control this API configures the maximal allowed current deviation between the set point and the actual current.
///
///=======
/// Remarks:
///=======
///   + Maximal allowed deviation between the set point and the actual current is 500mA.
///   + If the value exceeds, the fault OR (out of range) is set after the debounce time elapses, but the output is not disabled. If the deviation again falls below the 500mA value, the fault is cleared again after the debounce time elapses. 
///   + For more information see |bds_out_po_getStatus|.
///   + This function should be called only once in the application.
///
///----------
/// FFI:
///----------
///This API can be used in trusted partitions . For untrusted partitions use |bds_out_poc_cfg_ffi|. See Freedom from Interference (FFI) concept for more details.
///  
///==================================================================		  			===================================================================================================
///Return value    								  									Description
///==================================================================		  			===================================================================================================
///0																					No error.
///1																					A parameter is invalid.
///
///==================================================================		   			===================================================================================================
///
///=======
///Code Example:
///=======
///============================================================================
///
///PROGRAM PLC_PRG
///
///  VAR
///  
///	Init_flag_u8:USINT:=0;
/// 
///  END_VAR
///  
///IF(Init_flag_u8=0) THEN (*To make api call once in application*)
///		
///	(* configure current control for output K73 *)
///	
///	bds_out_poc_cfg(bds_out_po_signal_te.K73, 100);
///  
///	Init_flag_u8:=1;
///  
///END_IF
///
///============================================================================
{attribute 'external_name' := 'cmp_rts_bds_out_poc_cfg'}
FUNCTION bds_out_poc_cfg : USINT
VAR_INPUT
	///The connector assigned signal name of the output.
	signal_e: UINT;
	///Allowed current deviation [mA].
	///   + Range:0 to 500
	iDeviation_u16: UINT;
END_VAR

END_FUNCTION

// I/O API/OUT/FFI_API/bds_out_poc_cfg_ffi
{attribute 'external_name' := 'cmp_rts_bds_out_poc_cfg_ffi'}
FUNCTION bds_out_poc_cfg_ffi : USINT
VAR_INPUT
	///The connector assigned signal name of the output.
	signal_e: UINT;
	///Allowed current deviation [mA].
	///   + Range:0 to 500
	iDeviation_u16: UINT;
END_VAR

END_FUNCTION

// I/O API/OUT/FFI_API/bds_out_poc_ffi
{attribute 'external_name' := 'cmp_rts_bds_out_poc_ffi'}
FUNCTION bds_out_poc_ffi : USINT
VAR_INPUT
	///The connector assigned signal name of the output.
	signal_e: UINT;
	///Set point [mA].
	///   + Range:0 to 4000
	iSet_u16: UINT;
END_VAR

END_FUNCTION

// I/O API/OUT_LEGACY/bds_out_po_cfg
///Configures the proportional output with current measurement as a proportional output with current control (POC).
///
///=======
/// Remarks:
///=======
///   + With the current control are further configurations possible:
///	   + Software dither, see |bds_out_poc_cfgDither|.
///	   + Deviation of actual current from the set point. (see |bds_out_poc_cfg|.)
///   + For more information see |bds_out_po_getStatus|.
///   + This function should be called only once in the application.
///
///----------
/// FFI:
///----------
///This API can be used in trusted partitions . For untrusted partitions use |bds_out_po_cfg_ffi|. See Freedom from Interference (FFI) concept for more details.
///   
///------
/// Info:
///------
///
///Only the proportional outputs with current measurement can be configured as POC.
///
///==================================================================		  			===================================================================================================
///Return value    								  									Description
///==================================================================		  			===================================================================================================
///0																					No error.
///1																					A parameter is invalid.
///2																					output is disabled.
///
///==================================================================		   			===================================================================================================
///
///=======
///Code Example:
///=======
///============================================================================
///
///PROGRAM PLC_PRG
///
///  VAR
///  
///	Init_flag_u8:USINT:=0;
/// 
///  END_VAR
///  
///IF(Init_flag_u8=0) THEN (*To make api call once in application*)
///		
///	(* configure  proportional output with current control (POC) *)
///	
///	bds_out_po_cfg(bds_out_po_signal_te.K73, STD_ON);
///	
///	Init_flag_u8:=1;
///  
///END_IF
///
///============================================================================
{attribute 'external_name' := 'cmp_rts_bds_out_po_cfg'}
FUNCTION bds_out_po_cfg : USINT
VAR_INPUT
	///The connector assigned signal name of the output.
	signal_e: UINT;
	///Configure closed loop control.
	///   + STD_OFF - Deactive closed loop control
	///   + STD_ON   - Active closed loop control
	cfgPOC_u8: USINT;
END_VAR

END_FUNCTION

// I/O API/OUT_LEGACY/bds_out_poc_cfgDither
///Configures the software dither of a proportional output with closed loop control.
///
///=======
/// Remarks:
///=======
///   + The dither frequencies are predefined (see example below) and its amplitude range is from  0 to 500mA.
///   + For more information see |bds_out_po_getStatus|.
///   + The structure member status_b16 holds the information regarding the configuration.
///   + This function should be called only once in the application.
/// 
///----------
/// FFI:
///----------
///This API can be used in trusted partitions  For untrusted partitions use |bds_out_poc_cfgDither_ffi|. See Freedom from Interference (FFI) concept for more details.
///  
///------
/// Info:
///------
///
///The function is only possible for proportional outputs which has been configured as closed loop control.
///
///==================================================================		  			===================================================================================================
///Return value    								  									Description
///==================================================================		  			===================================================================================================
///0																					No error.
///1																					A parameter is invalid.
///2																					Wrong period for dither function.
///3																					Wrong dither frequency.
///
///==================================================================		   			===================================================================================================
///
///=======
///Code Example:
///=======
///============================================================================
///
///PROGRAM PLC_PRG
///
///VAR
///
///	Init_flag_u8:USINT:=0;
///
///END_VAR
///  
///IF(Init_flag_u8=0) THEN (*To make api call once in application*)
///			
///	(* configure the software dither output K73 *)
///	
///	bds_out_poc_cfgDither(bds_out_po_signal_te.K73, fDither_100Hz_DU8, 250);
///  
///	Init_flag_u8:=1;
///  
///END_IF
///
///
///============================================================================
{attribute 'external_name' := 'cmp_rts_bds_out_poc_cfgDither'}
FUNCTION bds_out_poc_cfgDither : USINT
VAR_INPUT
	///The connector assigned signal name of the output.
	signal_e: UINT;
	///Frequency [Hz]
	///
	///   + Range:Predefined values.
	frequency_u8: USINT;
	///Amplitude [mA]
	///
	///   + Range:0 to 500
	amplitude_u16: UINT;
END_VAR

END_FUNCTION

// I/O API/OUT/FFI_API/bds_out_poc_cfgDither_ffi
{attribute 'external_name' := 'cmp_rts_bds_out_poc_cfgDither_ffi'}
FUNCTION bds_out_poc_cfgDither_ffi : USINT
VAR_INPUT
	///The connector assigned signal name of the output.
	signal_e: UINT;
	///Frequency [Hz]
	///
	///   + Range:Predefined values.
	frequency_u8: USINT;
	///Amplitude [mA]
	///
	///   + Range:0 to 500
	amplitude_u16: UINT;
END_VAR

END_FUNCTION

// I/O API/OUT/FFI_API/bds_out_po_cfg_ffi
{attribute 'external_name' := 'cmp_rts_bds_out_po_cfg_ffi'}
FUNCTION bds_out_po_cfg_ffi : USINT
VAR_INPUT
	///The connector assigned signal name of the output.
	signal_e: UINT;
	///Configure closed loop control.
	///   + STD_OFF - Deactive closed loop control
	///   + STD_ON   - Active closed loop control
	cfgPOC_u8: USINT;
END_VAR

END_FUNCTION

// I/O API/IN legacy/API/bds_in_aic_getStatus
///Provides the status of the input.
///
///=======
/// Remarks:
///=======
///    + For information about the signal acquisition see Analog voltage aquisition.
///    + The status data provides all the relevant information regarding current input. See the example below.
///	    + The structure member status_b16 provides the information regarding the currently used configuration (also see  |bds_in_aic_cfg|) and the shunt status of the DSM frequency input.
///	    + Part of the status data also denotes the fault status of every DFC (e.g., stDFC_SCB_u16).  See  the topic Diagnostic Fault Check. 
///	    + With the macros (e.g., bds_dsm_DFC_ldf) defined in bds_dsm_api.h the respective bit fields of the fault status can be read.
///
///
///----------
/// FFI:
///----------
///This API can be used in trusted partitions only. See Freedom from Interference (FFI) concept for more details.
///
///==================================================================		  			===================================================================================================
///Return value    								  									Description
///==================================================================		  			===================================================================================================
///0																					No error
///1																					Invalid parameter
///
///==================================================================		   			===================================================================================================
///
///
///=======
///Code Example:
///=======
///============================================================================
///
///PROGRAM PLC_PRG
///
///  VAR
///  
///	Init_flag_u8:USINT:=0;
/// 
///  END_VAR
///  
///IF(Init_flag_u8=0) THEN (*To make api call once in application*)
///
///	(* As a precondition IN_CI_FI1 (K54_VI) must be switched once to a low resistance value *)
///	
///	bds_sys_do(bds_sys_do_signal_te.SHUNT1_EN, STD_ACTIVE);
///	
///	Init_flag_u8:=1;
///  
///END_IF
///
///PROGRAM appl_10ms_task
///  VAR
///  
///    stK54_s: bds_in_aic_ts;
///	
///    ldf_u8: USINT := 16#00;
///  END_VAR
///
///  (* get the status of input K54_VI *)
///
///  bds_in_aic_getStatus(bds_in_fi_signal_te.K54_VI, ADR(stK54_s));
///
///  (* get last debounced fault *)
///  
///  ldf_u8 = bds_dsm_DFC_ldf(stK54_s.stDFC_SCB_u16);
///END
///
///============================================================================
{attribute 'external_name' := 'cmp_rts_bds_in_aic_getStatus'}
FUNCTION bds_in_aic_getStatus : USINT
VAR_INPUT
	///The signal name that is assigned to the respective pin configured as current input
	signal_e: UINT;
	///Storage address of the data
	data_ps: POINTER TO bds_in_aic_ts;
END_VAR

END_FUNCTION

// I/O API/IN legacy/API/bds_in_aic_cfg
///Configures the diagnosis thresholds voltages of the input.
///
///=======
/// Remarks:
///=======
///   + The diagnosis is only possible after the configuration of the diagnosis thresholds. 
///	   + Depending on the configuration, the diagnosis threshold range for the configurable inputs can be from 150 to 4850 or 150 to 19850 or 150 to 39850mV.
///	   + The diagnosis threshold range for the fixed inputs ranges is from 150 to 29850mV.
///   + For more information see |bds_in_aiv_getStatus|.
///   + This function should be called only once in the application.
///
///----------
/// FFI:
///----------
///This API can be used in trusted partitions only. See Freedom from Interference (FFI) concept for more details.
///	
///==================================================================		  			===================================================================================================
///Return value    								  									Description
///==================================================================		  			===================================================================================================
///0																					No error
///1																					Invalid parameter
///2																					Function call was erroneous
///
///==================================================================		   			===================================================================================================
///
///=======
///Code Example:
///=======
///============================================================================
///
///PROGRAM PLC_PRG
///  VAR
///  
///	Init_flag_u8:USINT:=0;
///	
///  END_VAR
///
///IF(Init_flag_u8=0) THEN (*To make api call once in application*)
///
///	(* configure diagnosis thresholds of input K54_VI *)
///	
///	bds_in_aic_cfg(bds_in_fi_signal_te.K54_VI, 21000, 3000);
///	
///	Init_flag_u8:=1;
///  
///END_IF
///
///============================================================================
{attribute 'external_name' := 'cmp_rts_bds_in_aic_cfg'}
FUNCTION bds_in_aic_cfg : USINT
VAR_INPUT
	///The signal name that is assigned to the respective pin configured as voltage input
	signal_e: UINT;
	///Higher diagnosis threshold in [mV].
	///
	///Range:
	///
	///Configurable inputs:
	///150 to 4850 / 150 to 19850 / 150 to 39850
	///
	///Fixed inputs:
	///150 to 29850
	///
	///Note:
	///upperThreshold_u16 > lowerThreshold_u16
	upperThreshold_u16: UINT;
	///Lower diagnosis threshold in [mV].
	///
	///Range:
	///
	///Configurable inputs:
	///150 to 4850 / 150 to 19850 / 150 to 39850
	///
	///Fixed inputs:
	///150 to 29850
	///
	///Note:
	///lowerThreshold_u16 < upperThreshold_u16
	lowerThreshold_u16: UINT;
END_VAR

END_FUNCTION

// I/O API/IN legacy/API/bds_in_aiv_getStatus
///Provides the status of the input.
///
///=======
/// Remarks:
///=======
///   + For information about the signal acquisition see Analog voltage aquisition.
///   + The status data provides all relevant information about the voltage input as shown in the example below.
///	   + One component of the status data is also the fault status of every DFC (e.g., stDFC_SCB_u16). (see topic Diagnostic Fault Check. )
///	   + Using the macros (e.g. bds_dsm_DFC_ldf) defined in bds_dsm_api.h, the bits corresponding  to the bit fields of the fault status can be read.
///
///
///----------
/// FFI:
///----------
///This API can be used in trusted partitions only. See Freedom from Interference (FFI) concept for more details.
///
///==================================================================		  			===================================================================================================
///Return value    								  									Description
///==================================================================		  			===================================================================================================
///0																					No error
///1																					Invalid parameter
///
///==================================================================		   			===================================================================================================
///
///=======
///Code Example:
///=======
///============================================================================
///
///PROGRAM appl_10ms_task
///  VAR
///  
///    stK59_s: bds_in_aiv_ts;
///	
///    ldf_u8: USINT := 16#00;
///  END_VAR
///
/// (* configure the status of input K59 *)
/// bds_in_aiv_getStatus(bds_in_aiv_signal_te.K59, ADR(stK59_s));
///
/// (* get last debounced fault *)
/// ldf_u8 := bds_dsm_DFC_ldf(stK59_s.stDFC_SCB_u16);
///END
///
///============================================================================
{attribute 'external_name' := 'cmp_rts_bds_in_aiv_getStatus'}
FUNCTION bds_in_aiv_getStatus : USINT
VAR_INPUT
	///The signal name that is assigned to the respective pin configured as voltage input
	signal_e: UINT;
	///Storage address of the data.
	data_ps: POINTER TO bds_in_aiv_ts;
END_VAR

END_FUNCTION

